// TIA Portal V20 export
Screen "Pop-up_OVERVIEW_LEGEND_Popup"  360x480
  ScreenItem "Background" at 0,0 size 360x480  Type=HmiRectangle
  ScreenItem "Textfeld_Legende" at 1,1 size 358x25  Type=HmiTextBox
  ScreenItem "Textfeld_2" at 10,148 size 140x20  Type=HmiTextBox
  ScreenItem "Textfeld_1" at 10,126 size 140x20  Type=HmiTextBox
  ScreenItem "Textfeld_3" at 10,37 size 140x20  Type=HmiTextBox
  ScreenItem "Textfeld_4" at 10,60 size 140x20  Type=HmiTextBox
  ScreenItem "Textfeld_5" at 10,82 size 140x20  Type=HmiTextBox
  ScreenItem "Textfeld_6" at 10,104 size 140x20  Type=HmiTextBox
  ScreenItem "Textfeld_9" at 155,126 size 200x20  Type=HmiTextBox
  ScreenItem "Textfeld_10" at 155,148 size 200x20  Type=HmiTextBox
  ScreenItem "Textfeld_11" at 155,37 size 110x20  Type=HmiTextBox
  ScreenItem "Textfeld_12" at 155,60 size 200x20  Type=HmiTextBox
  ScreenItem "Textfeld_13" at 155,82 size 200x20  Type=HmiTextBox
  ScreenItem "Textfeld_14" at 155,104 size 200x20  Type=HmiTextBox
  ScreenItem "Cancel Mode" at 269,1 size 90x60  Type=HmiButton
  ScreenItem "Textfeld_7" at 10,207 size 335x54  Type=HmiTextBox
  ScreenItem "Textfeld_8" at 10,170 size 140x20  Type=HmiTextBox
  ScreenItem "Textfeld_15" at 154,163 size 200x36  Type=HmiTextBox
  ScreenItem "Linie_1" at 10,270 size 340x0  Type=HmiLine
  ScreenItem "Linie_2" at 10,271 size 340x0  Type=HmiLine
  ScreenItem "Textfeld_Legende_2" at 10,281 size 340x20  Type=HmiTextBox
  ScreenItem "Textfeld_16" at 10,309 size 345x36  Type=HmiTextBox
  ScreenItem "Textfeld_17" at 227,347 size 35x20  Type=HmiTextBox
  ScreenItem "Textfeld_18" at 308,347 size 45x20  Type=HmiTextBox
  ScreenItem "Textfeld_20" at 269,346 size 32x20  Type=HmiTextBox
  ScreenItem "Textfeld_19" at 183,347 size 32x20  Type=HmiTextBox
  ScreenItem "V_01" at 198,368 size 3x11  Type=HmiRectangle
  ScreenItem "H_01" at 191,379 size 17x3  Type=HmiRectangle
  ScreenItem "Textfeld_21" at 10,347 size 168x20  Type=HmiTextBox
  ScreenItem "Textfeld_22" at 10,380 size 330x20  Type=HmiTextBox
  ScreenItem "Textfeld_23" at 19,400 size 25x18  Type=HmiTextBox
  ScreenItem "Textfeld_24" at 127,400 size 25x18  Type=HmiTextBox
  ScreenItem "Textfeld_25" at 234,400 size 25x18  Type=HmiTextBox
  ScreenItem "Textfeld_26" at 50,399 size 75x20  Type=HmiTextBox
  ScreenItem "Textfeld_27" at 157,400 size 75x20  Type=HmiTextBox
  ScreenItem "Textfeld_28" at 264,400 size 75x20  Type=HmiTextBox
  ScreenItem "Textfeld_29" at 10,422 size 345x52  Type=HmiTextBox
